// TwinCAT 3 PLC project Training
// ProgramVersion: 3.1.4026.17
// libraries:
//   LCLS General, * (SLAC)
//   LCLS_Tc_DevAbs, * (SLAC - LCLS)
//   LCLS_Tc_Motion, * (SLAC - LCLS)
//   Tc2_EtherCAT, * (Beckhoff Automation GmbH)
//   Tc2_MC2, * (Beckhoff Automation GmbH)
//   Tc2_Standard, * (Beckhoff Automation GmbH)
//   Tc2_System, * (Beckhoff Automation GmbH)
// project tree:
//   DUTs/ E_AxisStates.TcDUT
//   GVLs/ GVL_Axes.TcGVL
//   / PlcTask.TcTTO
//   POUs/ PRG_SM.TcPOU, PRG_PTP.TcPOU
// real-time tasks:
//   TASK PlcTask: cycle T#10ms, priority 20, ADS port 350
// motion (NC):
//   TASK NC-Task 1 SAF: cycle T#2ms, priority 4, ADS port 501
//   TASK NC-Task 1 SVB: cycle T#10ms, priority 8, ADS port 511
//   AXIS HT23 (id 1)
//     Dynamic: AccelerationMaximum=10, DecelerationMaximum=10, Acceleration=10, Deceleration=10, Jerk=149.9985
//     Velo: RefSearch=0.33333, RefSync=0.33333, SlowManual=1.66665, FastManual=9.9999, Fast=33.333, Maximum=2
//     OtherSettings: AllowMotionCmdToSlave=true
//     encoder EncType=1
//       EncPara: ScaleFactorNumerator=4, ScaleFactorDenominator=1048576
//     drive DrvType=5
//       Analog: VeloReferenz=36.6663, TorqueSetpointScale=10, ScaleFactorActTorque=0.1
//       TimeComp: TaskDelayCycles=1
//     controller CtrType=1
//       CtrPara: PriorControlFactor=1
//         Observer: BandWidth=20
//   AXIS SO23HS (id 2)
//     OtherSettings: AllowMotionCmdToSlave=true
//     encoder EncType=1
//     drive DrvType=5
//       Analog: TorqueSetpointScale=10, ScaleFactorActTorque=0.1
//       TimeComp: TaskDelayCycles=1
//     controller CtrType=1
//       CtrPara: PriorControlFactor=1
//         Observer: BandWidth=20
// I/O:
//   DEVICE Device 1 (EtherCAT), AmsNetId 192.168.0.4.2.1
//     Term 1 (EK1101) [EK1101 EtherCAT Coupler (2A E-Bus, ID switch)]
//       Term 2 (EL5042) [EL5042 2Ch. BiSS-C Encoder]
//       Term 3 (EL7062) [EL7062-0000 2Ch. Stepper motor output stage (48V, 3A)]
//         startup 32785:27 := 4D420000 // DRV Motor Settings Ch.1 / Motor speed limitation
//         startup 28688:3 := 08 // DRV Outputs Ch.1 / Modes of operation
//         startup 28688:16 := FF7F // DRV Outputs Ch.1 / Positive torque limit value
//         startup 28688:17 := FF7F // DRV Outputs Ch.1 / Negative torque limit value
//         startup 32784:87 := 64 // DRV Amplifier Settings Ch.1 / Position loop velocity feed forward gain
//         startup 32784:109 := 64000000 // DRV Amplifier Settings Ch.1 / Torque feed forward gain
//         startup 32785:52 := B80B0000 // DRV Motor Settings Ch.1 / Configured motor current
//         startup 32784:19 := 3100 // DRV Amplifier Settings Ch.1 / Current loop proportional gain
//         startup 32784:18 := 1E00 // DRV Amplifier Settings Ch.1 / Current loop integral time
//         startup 32784:21 := 75000000 // DRV Amplifier Settings Ch.1 / Velocity loop proportional gain
//         startup 32784:20 := 96000000 // DRV Amplifier Settings Ch.1 / Velocity loop integral time
//       Term 4 (EL9011) [EL9011 End Terminal]
// variable links:
//   (this object) <-> NC-Task 1 SAF/Axes/HT23
//     PlcTask Inputs/GVL_Axes.Axes[1].NcToPlc <-> Outputs/ToPlc
//     PlcTask Outputs/GVL_Axes.Axes[1].PlcToNc <-> Inputs/FromPlc
//   (this object) <-> NC-Task 1 SAF/Axes/SO23HS
//     PlcTask Inputs/GVL_Axes.Axes[2].NcToPlc <-> Outputs/ToPlc
//     PlcTask Outputs/GVL_Axes.Axes[2].PlcToNc <-> Inputs/FromPlc

CONFIGURATION Training
    RESOURCE PLC ON TwinCAT3
        TASK PlcTask(INTERVAL := T#10ms, PRIORITY := 20);
        PROGRAM PRG_PTP WITH PlcTask : PRG_PTP;
    END_RESOURCE
END_CONFIGURATION

// ---- DUTs/E_AxisStates.TcDUT
{attribute 'qualified_only'}
{attribute 'strict'}
{attribute 'to_string'}
TYPE E_AxisStates :
(
    UNKNOWN := 0, // UNKNOWN must be in slot 0 or the FB breaks
    OUT := 1,
    YAG := 2,
    TT := 3
) UINT;
END_TYPE

// ---- GVLs/GVL_Axes.TcGVL
{attribute 'qualified_only'}
VAR_GLOBAL
    Axes :  ARRAY[1..4] OF AXIS_REF;
END_VAR

// ---- POUs/PRG_PTP.TcPOU
PROGRAM PRG_PTP
VAR
    fbPersistentDataStorage : LCLS_Tc_DevAbs.FB_PersistentDataStorage;
	{attribute 'pytmc' := '
		axis-link: GVL_Axes.Axes[1]
		pv: TST:MOTION:PTP
	'}
   	fbPtp : FB_MotionStageNC(	
		sName := 'PTP',
        AxisRef := GVL_Axes.Axes[1],
        iPersistentDataStorage := fbPersistentDataStorage
	) ;
	bFirstScan: BOOL := TRUE;
END_VAR

IF bFirstScan THEN
    fbPtp.SetModeEnableLimits(
        LimBackward := TRUE,
        LimForward := TRUE,
        HomeEnable  := FALSE,
        BrakeMode   := E_StageBrakeMode.IF_ENABLED,
        EnableMode  := E_StageEnableMode.DURING_MOTION,
        HomeMode    := 1,
        UserEnable  := TRUE,
        HardwareEnable := TRUE
    );
    fbPtp.SetVelocity(
        Velocity     := 1.0
    );
    bFirstScan := FALSE;
END_IF

fbPtp();
fbPersistentDataStorage();

END_PROGRAM

// ---- POUs/PRG_SM.TcPOU
PROGRAM PRG_SM
VAR
fbPersistentDataStorage : LCLS_Tc_DevAbs.FB_PersistentDataStorage;
	{attribute 'pytmc' := '
		pv: TST:MOTION
		io: io
		axis-link: GVL_Axes.Axes[1], GVL_Axes.Axes[2]
		expand-names: M1, M2
	'}	
    afbMotorsNC	: ARRAY[1..MotionConstants.MAX_STATE_MOTORS] OF FB_MotionStageNC[
		(AxisRef := GVL_Axes.Axes[1],  iPersistentDataStorage := fbPersistentDataStorage,  sName := 'M1'),
		(AxisRef := GVL_Axes.Axes[2],  iPersistentDataStorage := fbPersistentDataStorage,  sName := 'M2')
	];
	{attribute 'pytmc' := '
		pv: TST:MOTION:STATE
		io: io
		expand-names: M1, M2
	'}
    astPositionState	:  ARRAY[1..MotionConstants.MAX_STATE_MOTORS] OF ARRAY[1..GeneralConstants.MAX_STATES] OF ST_PositionState;
    aiMotionStage     	:  ARRAY[1..MotionConstants.MAX_STATE_MOTORS] OF I_MotionStage
                        := [afbMotorsNC [1], afbMotorsNC[2]];
    {attribute 'pytmc' := '
          pv: TST:MOTION:STATE:SET
          io: io
    '}
    eEnumSet          	: E_AxisStates;
    {attribute 'pytmc' := '
          pv: TST:MOTION:STATE:GET
          io: i
    '}
    eEnumGet          	: E_AxisStates;
	
    stDefault : ST_PositionState := (
        fDelta := 0.5,
        bMoveOk := TRUE,
        bValid := TRUE
    );
    fbStateConfigurator : FB_StateConfigurator(
        stDefault:= stDefault,
        bSetDefault:=TRUE
    );
//Configurators
    afbStateConfig : ARRAY[1..MotionConstants.MAX_STATE_MOTORS * GeneralConstants.MAX_STATES]
                       OF FB_StateConfigurator[
        // Motor 1
        (stPositionState := astPositionState[1][E_State.OUT],      stDefault := stDefault, bSetDefault:= TRUE, sName := 'OUT',      fPosition := 100.0),
        (stPositionState := astPositionState[1][E_State.TARGET1A], stDefault := stDefault, bSetDefault:= TRUE, sName := 'TARGET1A', fPosition := 200.0),
        (stPositionState := astPositionState[1][E_State.TARGET1B], stDefault := stDefault, bSetDefault:= TRUE, sName := 'TARGET1B', fPosition := 300.0),
        (stPositionState := astPositionState[1][E_State.TARGET1C], stDefault := stDefault, bSetDefault:= TRUE, sName := 'TARGET1C', fPosition := 400.0),
        // Motor 2
        (stPositionState := astPositionState[2][E_State.OUT],      stDefault := stDefault, bSetDefault:= TRUE, sName := 'OUT',            fPosition := 100.0),
        (stPositionState := astPositionState[2][E_State.TARGET1A], stDefault := stDefault, bSetDefault:= TRUE, sName := 'TARGET1A',  fPosition := 200.0),
        (stPositionState := astPositionState[2][E_State.TARGET1B], stDefault := stDefault, bSetDefault:= TRUE, sName := 'TARGET1B',  fPosition := 300.0),
        (stPositionState := astPositionState[2][E_State.TARGET1C], stDefault := stDefault, bSetDefault:= TRUE, sName := 'TARGET1C',  fPosition := 400.0)
    ];
    {attribute 'pytmc' := 'pv: TST:MOTION'}
    fbPositionStateND : FB_PositionStateND(
        aiMotionStage    := aiMotionStage,
        astPositionState := astPositionState,
		nActiveMotorCount := 2,
        eEnumSet         := eEnumSet,
        eEnumGet         := eEnumGet
    );
    bFirstScan : BOOL := TRUE;
	rtReady: R_TRIG;
    i    : INT;
    nCfg : INT;
END_VAR

IF bFirstScan THEN
	FOR i := 1 TO 3 DO
		afbMotorsNC[i].SetModeEnableLimits(
			LimBackward    := TRUE,
			LimForward     := TRUE,
			HomeEnable     := FALSE,
			BrakeMode      := E_StageBrakeMode.IF_ENABLED,
			EnableMode     := E_StageEnableMode.DURING_MOTION,
			HomeMode       := 1,
			UserEnable     := TRUE,
			HardwareEnable := TRUE
		);
		// Motion parameters live on the drive layer, not the state.
		afbMotorsNC[i].SetMotionParam(
			Velocity     := 25.0,
			Acceleration := 250.0,
			Deceleration := 250.0,
			Jerk         := 2500.0
		);
        afbMotorsNC[i].RestoreMotionParams:= FALSE;
	END_FOR
    bFirstScan := FALSE;
END_IF

// Configure states : called every cycle. One configurator per (motor, state)
// pair, each bound to its own stPositionState reference at init.
FOR nCfg := 1 TO MotionConstants.MAX_STATE_MOTORS * GeneralConstants.MAX_STATES DO
    afbStateConfig[nCfg]();
END_FOR

fbPositionStateND();
fbPersistentDataStorage();
FOR i := 1 TO 2 DO
	afbMotorsNC[i]();	
END_FOR

END_PROGRAM
